(* ================================================================= *)
(*  类型名称：ST_Manual                                          *)
(*  功能描述：手动与示教状态 (FB_1006 写)                                *)
(*  版本号：V1.0.0 (2026-10-24, DJ-2026-005 新设计)                    *)
(*  依据：接口文档_INT.md                                              *)
(* ================================================================= *)

TYPE ST_Manual
STRUCT
    bJogLockZ               : BOOL;     // Z 轴点动禁止
    bJogLockX1              : BOOL;     // X1 轴点动禁止
    bJogLockX2              : BOOL;     // X2 轴点动禁止
    abForce                 : ARRAY[1..21] OF BOOL;     // 输送强制位 (已按条件放行), 下标 = 位置 + 1
    bTeachWrite             : ARRAY[1..6] OF BOOL;      // 示教写入脉冲
    bGripOpenCmd            : BOOL;     // 手动夹爪松开命令
    bLiftUpCmd              : BOOL;     // 手动升降缸上升命令
    bLiftDownCmd            : BOOL;     // 手动升降缸下降命令
    arrTrig                 : ARRAY[1..2] OF BOOL;      // 报警触发 (保留)
END_STRUCT
END_TYPE
